// TIA Portal V21 export
// export: Created 2026-11-11T00:47:10.3131934Z, ExportSetting WithDefaults, DisplayName Totally Integrated Automation Portal, DisplayVersion V21 Update 3, DisplayName STEP 7 Professional, DisplayVersion V21 Update 3, DisplayName STEP 7 Safety, DisplayVersion V21, DisplayName Tech WebApplication, DisplayVersion V21, DisplayName WinCC Basic/Comfort/Advanced, DisplayVersion V21 Update 3, DisplayName WinCC Unified, DisplayVersion V21 Update 3
FUNCTION_BLOCK "FB_Fbd_Put"   // FB345, FBD
{ S7_Optimized_Access := 'FALSE' }
VERSION : 0.1
// stored: AutoNumber true, IsIECCheckEnabled false, SetENOAutomatically false, UDAEnableTagReadback false
   VAR_INPUT
      req : Bool;
      id : Word;
   END_VAR
   VAR_OUTPUT
      done : Bool;
      err : Bool;
      status : Word;
   END_VAR
   VAR_IN_OUT
      addr1 : Remote;
      addr2 : Remote;
      addr3 : Remote;
      addr4 : Remote;
   END_VAR
   VAR
      inst { S7_SetPoint := 'True'} : PUT;
   END_VAR
   VAR_TEMP
      rd1 : Array[0..9] of Byte;
      rd2 : Array[0..9] of Byte;
      rd3 : Array[0..9] of Byte;
      rd4 : Array[0..9] of Byte;
   END_VAR
BEGIN

REGION Network 1: PUT
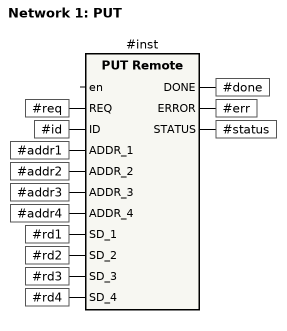
   #inst(REQ := #req,   // PUT
         ID := #id,
         ADDR_1 := #addr1,
         ADDR_2 := #addr2,
         ADDR_3 := #addr3,
         ADDR_4 := #addr4,
         SD_1 := #rd1,
         SD_2 := #rd2,
         SD_3 := #rd3,
         SD_4 := #rd4,
         DONE => #done,
         ERROR => #err,
         STATUS => #status);
END_REGION
END_FUNCTION_BLOCK
